//{attribute 'qualified_only'}
VAR_GLOBAL
	fbAnybus	: FB_Anybus_Interface;	//CIP <-> Siemens exchange, called in MAIN
	fbSim		: FB_Siemens_Sim;		//Siemens simulator, commissioning only
	bSimEnable	: BOOL;					//TRUE: fbSim replaces the gateway inputs
	arSimRaw	: ARRAY[0..127] OF BYTE;
	bQueueCleared	: BOOL;				//the persistent CIP queue is cleared once after PLC start
	fbBridge	: FB_CIP_Siemens;		//Siemens order -> FB_CIP, CIP state -> Siemens
	bBridgeEnable	: BOOL;				//FALSE: CIP runs from HMI only, stStatus is left alone
END_VAR

(* stored: Version 1.1.0.1, ProductVersion 3.1.4026.20
   GVL g_Anybus: Id {e0092543-9a36-4da0-b8be-76804fae3bd9} *)
